FUNCTION_BLOCK FB_STOEBERSDS_MC_AxisMoveManual
(*

The function block used to manual control of axis.

Constructor: 		Patryk Panylo
Company:		E. Riexinger GmbH
Date:			22.09.2015
Version:			1.00

Date:			Revision:		Who:				Comment
dd.mm.yyyy		x.xx			Initials			comment

*)
VAR_INPUT
	(* Input variables / Eingang Variablen *)
	bEnable						:BOOL;						(* Signal FB enable *)
	etMachineMode				:ET_MachineMode;			(* Machine mode *)
	etMachineState				:ET_MachineState;			(* Machine state *)
	bCtrlEnabled					:BOOL;						(* Controller enabled *)
	bReset						:BOOL;						(* Reset *)
	bMovePlus					:BOOL;						(* Move in plus direction *)
	bMoveMinus					:BOOL;						(* Move in minus direction *)
	lrTipDistance					:LREAL;						(* Relative distance for movements *)
	bLimitMax					:BOOL;						(* Limit max *)
	bLimitMin					:BOOL;						(* Limit min *)
	bPlusRelease				:BOOL;						(* Plus move release *)
	bMinusRelease				:BOOL;						(* Minus move release *)
	lrVelocity						:LREAL;						(* Target velocity *)
	lrAcceleration					:LREAL;						(* Value of the acceleration (always positive) *)
	lrDeceleration				:LREAL;						(* Value of deceleration (always positive) *)
	lrJerk						:LREAL;						(* Value of jerk (always positive) *)
	tControllerOff					:TIME := t#60s;				(* Time to switch controller off *)
END_VAR
VAR_OUTPUT
	(* Output variables / Ausgang Variablen *)
	bMoving						:BOOL;						(* Axis moving *)
	bControllerOff					:BOOL;						(* Switch controller off *)
	bBusy						:BOOL;						(* Program busy *)
	bError						:BOOL;						(* Program error *)
	udnErrorNo					:UDINT;						(* Error number *)
END_VAR
VAR_IN_OUT
	bHomeCompleted				:BOOL;						(* Home completed *)
	Axis							:ST_AXIS_REF;					(* The AXIS_REF data type  is an interface between the PLC and the NC and contains axis information *)
END_VAR
VAR
	(* Enummerations *)

	(* Variables *)
	bFirstTime					:BOOL;

	(* References *)

	(* Interfaces *)

	(* Instances *)
	fbJog						:FB_STOEBERSDS_MC_Jog;					(* The function block is used to manual control an axis *)
	fbTipPlus					:FB_SignalWatchdog;
	fbTipMinus					:FB_SignalWatchdog;
	rtMovePlus					:R_TRIG;
	rtMoveMinus					:R_TRIG;
END_VAR


IF NOT bEnable							(* Signal FB enable *)
THEN
	fbJog(
		bEnable := FALSE,
		bJogForward := FALSE,
		bJogBackwards := FALSE,
		Axis := Axis,
		bActive => bMoving				(* Axis moving *)
	);

	fbTipPlus(
		bEnable := FALSE,
		tWatchdog := tControllerOff
	);

	fbTipMinus(
		bEnable := FALSE,
		tWatchdog := tControllerOff
	);

	bControllerOff := FALSE;

	bFirstTime := FALSE;

	RETURN;
END_IF

IF NOT bFirstTime
THEN

	bFirstTime := TRUE;
END_IF

IF bReset
     AND bError
THEN
	fbJog(
		bEnable := FALSE,
		bJogForward := FALSE,
		bJogBackwards := FALSE,
		Axis := Axis,
		bActive => bMoving				(* Axis moving *)
	);
END_IF;

A_SetLimits();

IF bCtrlEnabled
    AND etMachineMode = ET_MachineMode_eManual
THEN
	rtMovePlus(CLK := bMovePlus);
	rtMoveMinus(CLK := bMoveMinus);

	IF NOT bMovePlus
	     AND NOT bMoveMinus
	THEN
		fbJog.bJogForward := FALSE;
		fbJog.bJogBackwards := FALSE;

	ELSIF bMovePlus
	             AND NOT bMoveMinus
	THEN
		fbJog.bJogForward := (lrTipDistance = 0 OR rtMovePlus.Q)
							    AND bPlusRelease AND NOT bLimitMax;
		fbJog.bJogBackwards := FALSE;
	
	ELSIF NOT bMovePlus
	     	    AND bMoveMinus
	THEN
		fbJog.bJogForward := FALSE;
		fbJog.bJogBackwards := (lrTipDistance = 0 OR rtMoveMinus.Q)
							          AND bMinusRelease AND NOT bLimitMin;
	
	END_IF;

	fbJog(
		bEnable := TRUE,
		etMode := SEL(lrTipDistance <> 0, ET_JogMode_MC_JOGMODE_STANDARD, ET_JogMode_MC_JOGMODE_INCHING),
		lrPosition := lrTipDistance,
		lrVelocity := lrVelocity,
		lrAcceleration := lrAcceleration,
		lrDeceleration := lrDeceleration,
		lrJerk := lrJerk,
		Axis := Axis,
		bActive => bMoving
	);

ELSE
	fbJog(
		bJogForward := FALSE,
		bJogBackwards := FALSE,
		Axis := Axis,
		bActive => bMoving				(* Axis moving *)
	);

END_IF

fbTipPlus(
	bEnable := etMachineMode = ET_MachineMode_eManual,
	bIn := bMovePlus
		  AND bPlusRelease
		  AND NOT bLimitMax,
	tWatchdog := tControllerOff
);

fbTipMinus(
	bEnable := etMachineMode = ET_MachineMode_eManual,
	bIn := bMoveMinus
		  AND bMinusRelease
		  AND NOT bLimitMin,
	tWatchdog := tControllerOff
);


bControllerOff := NOT (fbTipPlus.bOut
			    	       OR fbTipMinus.bOut)
			    AND etMachineMode = ET_MachineMode_eManual;

IF bMoving
THEN
	bHomeCompleted := FALSE;
END_IF;

bError := fbJog.bError;

ACTION A_SetLimits:
;
END_ACTION

END_FUNCTION_BLOCK

(* stored: Version 1.1.0.1, ProductVersion 3.1.4024.15
   POU FB_STOEBERSDS_MC_AxisMoveManual: Id {dc454482-85a8-482b-9e38-77799a196d2f}, SpecialFunc None
   Action A_SetLimits: Id {9a71e1a8-b875-4b33-b962-a1078bbecfb4} *)
